TYPE "ST_PressDemoStationCfg"
VERSION : 0.1
   STRUCT
      SchemaVersion : UInt := 1;
      RequireTwoHandStart : Bool := TRUE;
   END_STRUCT;

END_TYPE

